RESOURCE RES0 : EMB_RES_ECO
  FBS
    FullInit : DPAC_FULLINIT;
    Sorting : Sorting(QI := TRUE);
    SeqInit : EVENTCHAINHEAD(NAME := 'SEQ_INIT');
  END_FBS
  EVENT_CONNECTIONS
    START.COLD TO FullInit.INIT;
    START.WARM TO FullInit.INIT;
    START.ONLINECHANGE TO FullInit.OC_RETRIGGER;
    FullInit.INITO TO SeqInit.INIT;
    FullInit.OC_DONE TO SeqInit.RETRIGGER;
    SeqInit.INITO TO SeqInit.TRIGGER;
    SeqInit.FINISHED TO Sorting.BB7E654A10914CAA;
  END_CONNECTIONS
END_RESOURCE
